///
///----------
/// FFI:
///----------
/// This API can be used in both trusted and untrusted partitions. See Freedom from Interference (FFI) concept for more details.
///
///------
///
///==================================================================		  			===================================================================================================
///Return value    								  									    Description
///==================================================================		  			===================================================================================================
///bds_outPwm_get_ts												                   The return structure containing;
///																							- Set current value in [mA]
///																							- Actual current measurement/current sensing of average of one PWM period in [mA]
///																							- Set value duty cycle in [permil]
///																							- Detailed diagnostic information OF the PWM output.
///																							- Function call status information (statusApi_e)
///
///==================================================================		   			===================================================================================================
///
///=======
///Code Example:
///=======
///============================================================================
///
/// PROGRAM appl_10ms_task
///
/// VAR
///
///     bds_outPwm_signal_e: bds_outPwm_signal_te; (* Declare the type for Pwm output signal*)
///
///     bds_outPwm_retGet_s: bds_outPwm_get_ts;    (* Declare the return structure of BDS-Function call*)
///
/// END_VAR
/// 
/// (* Initialize the signal value*)
///
/// bds_outPwm_signal_e := bds_outPwm_signal_te.bds_outPwm_K09_E;
/// 
/// (* Call BDS-Function to get the status of the output*)
///
/// bds_outPwm_retGet_s := bds_outPwm_get(bds_outPwm_signal_e);
/// 
/// (* Check return state of BDS-Function call*)
///
/// IF bds_outCmn_ok_E = bds_outPwm_retGet_s.statusApi_e THEN
///
///     (* Call successful, signal is valid*)
///
///     (* Status of output is updated successfully*)
///
/// ELSE
///
///     (* Handle error*)
///
/// END_IF;
///
/// END_PROGRAM
///
///============================================================================
{attribute 'external_name' := 'cmp_rts_bds_outPwm_get'}
FUNCTION bds_outPwm_get : bds_outPwm_get_ts
VAR_INPUT
	///The connector assigned signaVl name of the output.
	signal_e: USINT;
END_VAR

END_FUNCTION

// I/O API/OUT/API/bds_outPwm_cfgPeriod
///The BODAS API-function configures the period of a PWM high side or low side output in [us].
///
///=======
/// Remarks:
///=======
/// FOR the "low power low side outputs" the period range is FROM FROM 300us upto 31000us.

/// For the "high power high side outputs" the period range is from 1000us upto 100000us and for the "high power low side outputs" 4000us upto 100000us and only multiples of 1000us is configurable.

/// Default value of period is 10000us.
///
///----------
/// FFI:
///----------
/// This API can be used in trusted partitions. For untrusted partitions use bds_outPwm_cfgPeriod_ffi. See Freedom from Interference (FFI) concept for more details.
///
///------
///
///==================================================================		  			===================================================================================================
///Return value    								  									    Description
///==================================================================		  			===================================================================================================
///bds_outPwm_cfgPeriod_ts														            The return structure containing the state information (statusApi_e)
///
///==================================================================		   			===================================================================================================
///
///=======
///Code Example:
///=======
///============================================================================
///
/// PROGRAM appl_10ms_task
///
/// VAR
///
///     bds_outPwm_signal_e: bds_outPwm_signal_te; (* Define the structure of Pwm output signal*)
///
///     bds_outPwm_retCfgPeriod_s: bds_outPwm_cfgPeriod_ts; (* Declare return structure for the function call*)
///
///     tiPerd_us_u32: UDINT := 1000; (* Define the period in microseconds*)
///
/// END_VAR
/// 
/// (* Assign the Pwm signal type*)
///
/// bds_outPwm_signal_e := bds_outPwm_signal_te.bds_outPwm_K09_E;
/// 
/// (* Call function to configure the period of a Pwm output*)
///
/// bds_outPwm_retCfgPeriod_s := bds_outPwm_cfgPeriod(bds_outPwm_signal_e, tiPerd_us_u32);
/// 
/// (* Check return state of the BDS-Function call*)
///
/// IF bds_outCmn_ok_E = bds_outPwm_retCfgPeriod_s.statusApi_e THEN
///
///     (* If the call was successful and the signal is valid*)
///
///     (* The period of the Pwm output has been configured successfully*)
///
/// ELSE
///
///     (* Error handling*)
///
/// END_IF;
///
/// END_PROGRAM
///============================================================================
{attribute 'external_name' := 'cmp_rts_bds_outPwm_cfgPeriod'}
FUNCTION bds_outPwm_cfgPeriod : bds_outPwm_cfgPeriod_ts
VAR_INPUT
	///The connector assigned signal name of the output.
	signal_e: USINT;
	///The connector assigned signal name of the output.
	tiPerd_us_u32: UDINT;
END_VAR

END_FUNCTION

// I/O API/OUT/API/bds_outPwm_rstErr
/// The BODAS API-function reset the diagnostics error and unlocks the PWM high side or low side output.
///=======
/// Remarks:
///=======
/// +After a fault, the output is locked but the set point is still valid. With the reset OF the error the output is also unlocked.

/// +After a hot short circuit, the unlocking of the power output is only possible after a reactivation time of 2s.

/// +It is possible to poll the status of the fault. If the error has been healed, then the output can be reset.

/// +For over current fault: After reset, the output has to be switched on again using the API bds_outPwm_setDutyCycle or bds_outPwm_setCurrent.

/// +For more information see topic Proportional outputs.


///----------
/// FFI:
///----------
/// This API can be used in trusted partitions. For untrusted partitions use bds_outPwm_rstErr_ffi. See Freedom from Interference (FFI) concept for more details.
///
///
///==================================================================		  			===================================================================================================
///Return value    								  									    Description
///==================================================================		  			===================================================================================================
///bds_outPwm_rstErr_ts													                The return structure containing the state information (statusApi_e)
///
///==================================================================		   			===================================================================================================
///
///=======
///Code Example:
///=======
///============================================================================
/// PROGRAM appl_10ms_task
///
/// VAR
///
///     bds_outPwm_signal_e: bds_outPwm_signal_te; (* Define the structure of Pwm output signal*)
///
///     bds_outPwm_retRstErr_s: bds_outPwm_rstErr_ts; (* Declare return structure for the function call
///
/// END_VAR
/// 
/// (* Assign the Pwm signal type*)
///
/// bds_outPwm_signal_e := bds_outPwm_signal_te.bds_outPwm_K09_E;
/// 
/// (* Call function to reset the Pwm output diagnostic error and unlock the Pwm output*)
///
/// bds_outPwm_retRstErr_s := bds_outPwm_rstErr(bds_outPwm_signal_e);
/// 
/// (* Check return state of the BDS-Function call*)
///
/// IF bds_outCmn_ok_E = bds_outPwm_retRstErr_s.statusApi_e THEN
///
///     (* If the call was successful and the signal is valid*)
///
///     (* The diagnostic error for the output has been reset and the output is unlocked*)
///
/// ELSE
///
///     (* Error handling*)
///
/// END_IF;
///
/// END_PROGRAM
///
///============================================================================
{attribute 'external_name' := 'cmp_rts_bds_outPwm_rstErr'}
FUNCTION bds_outPwm_rstErr : bds_outPwm_rstErr_ts
VAR_INPUT
	///The connector assigned signal name of the output.
	signal_e: USINT;
END_VAR

END_FUNCTION

// I/O API/OUT/API/bds_outPwm_setCurrent
///The BODAS API-function sets the current for the PWM high side or low side output which is configured as closed loop current control mode.
///
///Set current range is from 0mA upto 3000mA/4000mA Current control upper limit depends on the used output, refer to RC27-18/40 - Outputs
///
///=======
/// Remarks:
///=======
///  + After a fault the output is locked but the set point is still valid.
///
///  + For more information see topic Proportional outputs.

///
///
///----------
/// FFI:
///----------
///This API can be used in trusted partitions . For untrusted partitions use |bds_out_do_getCurrent_ffi|. See Freedom from Interference (FFI) concept for more details.
///
///---------
/// Info
///---------
/// It is mandatory that the proportional output is configured as proportional output with closed loop current control mode, refer to bds_outPwm_cfgMode.

///---------
/// Attention
/// ---------
/// It is possible to poll the status of the fault. If the error has been healed, then the output can be unlocked by calling THIS API-FUNCTION.
///
/// After a hot short circuit and over current the unlock of the high power output is only possible after a reactivation wait time of 2s, refer to bit in status bds_outCmn_statusDiag_tb.

///==================================================================		  			===================================================================================================
///Return value    								  									    Description
///==================================================================		  			===================================================================================================
/// bds_outPwm_setCurrent_ts															The return structure containing the state information (statusApi_e)
///
///==================================================================		   			===================================================================================================
///
///=======
///Code Example:
///=======
///============================================================================
///
/// PROGRAM appl_10ms_task
///
/// VAR
///
///  bds_outPwm_signal_e: bds_outPwm_signal_te; (* Structure of PWM output signal*)
///
///  bds_outPwm_cfgMode_e: bds_outPwm_cfgMode_te; (* Output mode structure*)
///
///  bds_outPwm_retSetCurrent_s: bds_outPwm_setCurrent_ts; (* Return structure for setting current*)
///
///  bds_outPwm_set_i_mA_u16: UINT := 500; (* Define the set-current in mA*)
///
/// END_VAR
///
////// bds_outPwm_signal_e := bds_outPwm_signal_te.bds_outPwm_K09_E;
/// 
/// (* Configure the output as closed loop control mode*)
///
/// bds_outPwm_cfgMode(bds_outPwm_signal_e, bds_outPwm_cfgMode_e);
/// 
/// (* Actuate the PWM output with set-current*)
///
/// bds_outPwm_retSetCurrent_s := bds_outPwm_setCurrent(bds_outPwm_signal_e, bds_outPwm_set_i_mA_u16);
/// 
/// (* Check the return state of the BDS-Function call*)
///
/// IF bds_outCmn_ok_E = bds_outPwm_retSetCurrent_s.statusApi_e THEN
///
///     (* If the call was successful and the signal is valid*)
///
///     (* The PWM output has been actuated to the requested set-current successfully*)
///
/// ELSE
///
///     (* Error handling*)
///
/// END_IF;
///
/// END_PROGRAM
///============================================================================
{attribute 'external_name' := 'cmp_rts_bds_outPwm_setCurrent'}
FUNCTION bds_outPwm_setCurrent : bds_outPwm_setCurrent_ts
VAR_INPUT
	///The connector assigned signal name of the output.
	signal_e: USINT;
	///Storage address of the value.
	///
	///   defining the set current value for a PWM output which is configured as closed loop control current with the resolution in [mA]
	i_mA_u16: UINT;
END_VAR

END_FUNCTION

// I/O API/OUT/API/bds_outPwm_cfgMode
///The BODAS API-function configures the PWM high side or low side output as closed loop current control mode.
///
///=======
/// Remarks:
///=======
///With the closed loop current control mode further configurations are possible:
///
/// Software dither, refer to bds_outPwm_cfgDither.
///
/// Allowed current deviation from the set point, refer to bds_outPwm_cfgDiagCurrentDe.
///
/// Gain PI-Controller values for regulation (Kp and Ki), refer to bds_outPwm_cfgClc.



///
///----------
/// FFI:
///----------
/// This API can be used in both trusted and untrusted partitions. See Freedom from Interference (FFI) concept for more details.
///
///------
/// Info
///------
/// Only the proportional outputs with "Current Measurement" can be configured as closed loop current control mode which means output can be actuated with set-current.
///
/// Default output is in Pwm mode which means output can only be actuated with duty-cycle

///
///==================================================================		  			===================================================================================================
///Return value    								  									    Description
///==================================================================		  			===================================================================================================
///bds_outPwm_cfgMode_ts													            The return structure containing the state information (statusApi_e)
///
///==================================================================		   			===================================================================================================
///
///=======
///Code Example:
///=======
///============================================================================
///
///PROGRAM appl_10ms_task
///
///
///VAR
///
///    bds_outPwm_signal_e: bds_outPwm_signal_te; (* Declare and define the structure of Pwm output signal*)
///
///    bds_outPwm_cfgMode_e: bds_outPwm_cfgMode_te; (* Declare and define the output mode structure*)
///
///    bds_outPwm_retCfgMode_s: bds_outPwm_cfgMode_ts; (* Declare the return structure of BDS-Function call*)
///
///END_VAR
///
///(* Assign the Pwm signal type*)
///
///bds_outPwm_signal_e := bds_outPwm_signal_te.bds_outPwm_K09_E;
///
///(* Set the output mode to closed loop current control*)
///
///bds_outPwm_cfgMode_e := bds_outMode_CLCC_E;
///
///(* Call function to configure the output as closed loop current control mode*)
///
///bds_outPwm_retCfgMode_s := bds_outPwm_cfgMode(bds_outPwm_signal_e, bds_outPwm_cfgMode_e);
///
///(* Check return state of the BDS-Function call*)
///
///IF bds_outCmn_ok_E = bds_outPwm_retCfgMode_s.statusApi_e THEN
///
///    (* If the call was successful and the signal is valid*)
///
///    (* Output has been configured as closed loop current control successfully*)
///ELSE
///
///    (* Error handling*)
///
///END_IF;
///
/// END_PROGRAM
///============================================================================
{attribute 'external_name' := 'cmp_rts_bds_outPwm_cfgMode'}
FUNCTION bds_outPwm_cfgMode : bds_outPwm_cfgMode_ts
VAR_INPUT
	///The connector assigned signal name of the output.
	signal_e: USINT;
	///The connector assigned signal name of the output.
	mode_e: bds_outPwm_cfgMode_te;
END_VAR

END_FUNCTION

// I/O API/OUT/API/bds_outPwm_cfgDither
///The BODAS API-function configure the dither frequency and amplitude for the PWM high side or low side output which is configured as closed loop current control mode.
///
///=======
/// Remarks:
///=======
///   + The dither frequencies are predefined (see bds_outPwm_cfgDither_te) and its amplitude range is from 0 to 500mA.
///
///   + Default value for dither frequency is 0 [Hz] and amplitude is 0 [mA] (means dither configuration is disabled).
/// 
///----------
/// FFI:
///----------
///This API can be used in trusted partitions. For untrusted partitions use bds_outPwm_cfgDither_ffi. See Freedom from Interference (FFI) concept for more details.
///  
///------
/// Info:
///------
///
///The function is only possible for proportional outputs which has been configured as closed loop current control mode and a period of 1ms (f = 1000 Hz), refer to Outputs PWM  RC27-18/40 - Outputs
///
///==================================================================		  			===================================================================================================
///Return value    								  										 Description
///==================================================================		  			===================================================================================================
///bds_outPwm_cfgDither_ts																bds_outPwm_cfgDither_ts															
///
///==================================================================		   			===================================================================================================
///
///=======
///Code Example:
///=======
///============================================================================
///
/// PROGRAM appl_10ms_task 
///
/// VAR
///
///     bds_outPwm_signal_e: bds_outPwm_signal_te; (* Structure of PWM output signal*)
///
///     bds_outPwm_cfgMode_e: bds_outPwm_cfgMode_te; (* Output mode structure*)
///
///     bds_outPwm_cfg_ditherParams_s: bds_outPwm_ditherParams_ts; (* Structure for dither parameters.*)
///
///     bds_outPwm_retCfgDither_s: bds_outPwm_cfgDither_ts; (* Return structure for the dither configuration function*)
///
///     tiPerd_us_u32: UDINT := 1000; (* Define the period in microseconds
///
/// END_VAR
/// 
/// (* Set the PWM signal type*)
///
/// bds_outPwm_signal_e := bds_outPwm_signal_te.bds_outPwm_K09_E;
/// 
/// (* Configure the output as closed loop control mode*)
///
/// bds_outPwm_cfgMode(bds_outPwm_signal_e, bds_outPwm_cfgMode_e);
/// 
/// (* Set dither frequency and amplitude*)
///
/// bds_outPwm_cfg_ditherParams_s.ditherFrq_Hz_e := bds_outPwm_dither_90_Hz_E;
///
/// bds_outPwm_cfg_ditherParams_s.ditherAmp_mA_u16 := 400;
/// 
/// (* Configure the period for PWM output*)
///
/// bds_outPwm_cfgPeriod(bds_outPwm_signal_e, tiPerd_us_u32);
/// 
/// (* Configure the dither frequency and amplitude*)
///
/// bds_outPwm_retCfgDither_s := bds_outPwm_cfgDither(bds_outPwm_signal_e, bds_outPwm_cfg_ditherParams_s);
/// 
/// (* Check return state of the BDS-Function call*)
///
/// IF bds_outCmn_ok_E = bds_outPwm_retCfgDither_s.statusApi_e THEN
///
///     (* If the call was successful and the signal is valid,*)
///
///     (* The dither frequency and amplitude for the PWM output have been configured successfully*)
///
/// ELSE
///
///     (* Error handling*)
///
/// END_IF;
///
/// END_PROGRAM
///
///============================================================================
{attribute 'external_name' := 'cmp_rts_bds_outPwm_cfgDither'}
FUNCTION bds_outPwm_cfgDither : bds_outPwm_cfgDither_ts
VAR_INPUT
	///defining the output signal for the PWM output
	signal_e: USINT;
	///Frequency [Hz]
	///
	///   + defining the control structure values for the dither frequency and amplitude values of the selected PWM output which is configured as Closed Loop Control Current
	ditherParams_s: bds_outPwm_ditherParams_ts;
END_VAR

END_FUNCTION

// I/O API/OUT/API/bds_outPwm_cfgDiagCurrentDe
/// The BODAS API-function sets the current deviation for the PWM high side or low side output which is configured as closed loop current control mode.
/// 
///
///=======
/// Remarks:
///=======
///
/// Maximal allowed deviation between the set point AND the actual current is 500mA.
///
/// Value of 0mA deviation means the current deviation monitoring is disabled.
///
///If the value exceeds, the fault OR (out of range) is set after the debounce time elapses, but the output is not switched OFF.
///
/// If the deviation falls below the set deviation value, the fault OR is cleared after the debounce time elapses. 
///
/// For more information see bds_outPwm_get.


 
///----------
/// FFI:
///----------
///This API can be used in trusted partitions. For untrusted partitions use bds_outPwm_cfgDiagCurrentDe_ffi. See Freedom from Interference (FFI) concept for more details.
///
///
///==================================================================		  			===================================================================================================
///Return value    								  									    Description
///==================================================================		  			===================================================================================================
///bds_outPwm_cfgDiagCurrentDe_ts														The return structure containing the state information (statusApi_e)
///
///==================================================================		   			===================================================================================================
///
///=======
///Code Example:
///=======
///============================================================================
///
///PROGRAM appl_10ms_task
///
///VAR
///
///    bds_outPwm_signal_e: bds_outPwm_signal_te; (* Structure of PWM output signal*)
///
///    bds_outPwm_cfgMode_e: bds_outPwm_cfgMode_te; (* Output mode structure*)
///
///    bds_outPwm_retCfgDiagCurrentDe_s: bds_outPwm_cfgDiagCurrentDe_ts; (* Return structure for configuring current deviation*)
///
///    bds_outPwm_cfg_iDe_mA_u16: UINT := 300; (* Define the set-deviation in mA*)
///
/// END_VAR
///
/// bds_outPwm_signal_e := bds_outPwm_signal_te.bds_outPwm_K09_E;
///
///(* Configure the output as closed loop control mode*)
///
///bds_outPwm_cfgMode(bds_outPwm_signal_e, bds_outPwm_cfgMode_e);
///
///(* Call function to configure the current deviation*)
///
///bds_outPwm_retCfgDiagCurrentDe_s := bds_outPwm_cfgDiagCurrentDe(bds_outPwm_signal_e, bds_outPwm_cfg_iDe_mA_u16);
///
///(* Check the return state of the BDS-Function call*)
///
///IF bds_outCmn_ok_E = bds_outPwm_retCfgDiagCurrentDe_s.statusApi_e THEN
///
///    (* If the call was successful and the signal is valid*)
///
///    (* The current deviation for the PWM output has been configured successfully*)
///
///ELSE
///
///    (* Error handling*)
//
///END_IF;
///
/// END_PROGRAM
///============================================================================
{attribute 'external_name' := 'cmp_rts_bds_outPwm_cfgDiagCurrentDe'}
FUNCTION bds_outPwm_cfgDiagCurrentDe : bds_outPwm_cfgDiagCurrentDe_ts
VAR_INPUT
	///The connector assigned signal name of the output.
	signal_e: USINT;
	/// defining the deviation current value for a PWM output which is configured as closed loop control current with the resolution in [mA]
	iDe_mA_u16: UINT;
END_VAR

END_FUNCTION

// I/O API/OUT/API/bds_outPwm_cfgClc
///The BODAS API-function configure closed loop control gain for the PWM high side or low side output which is configured as closed loop current control mode.
///
///=======
/// Remarks:
///=======
///   +Range Kp factor [0...2000] and set default value is 100.
///
///	  +Range Ki factor [0...500] and set default value is 25.
///
///----------
/// FFI:
///----------
/// This API can be used in trusted partitions. For untrusted partitions use bds_outPwm_cfgClc_ffi. See Freedom from Interference (FFI) concept for more details.
///   
///==================================================================		  			===================================================================================================
///Return value    								  									     Description
///==================================================================		  			===================================================================================================
///bds_outPwm_cfgClc_ts																	The return structure containing the state information (statusApi_e)																		
///
///==================================================================		   			===================================================================================================
///
///=======
///Code Example:
///=======
///============================================================================
///
/// PROGRAM appl_10ms_task
///
/// VAR
///
///     bds_outClcC_signal_e: bds_outPwm_signal_te; (* Structure of PWM output signal*)
///
///     bds_outPwm_cfgMode_e: bds_outPwm_cfgMode_te; (* Output mode structure*)
///
///     bds_outPwm_cfg_clcParams_s: bds_outPwm_clcParams_ts; (* Structure for closed loop control gain*)
///
///     bds_outPwm_retCfgClc_s: bds_outPwm_cfgClc_ts; (* Return structure of BDS-Function call*)
///
/// END_VAR
/// 
/// (* Set the PWM signal type*)
///
/// bds_outClcC_signal_e := bds_outPwm_signal_te.bds_outPwm_K09_E;
/// 
/// (* Configure the output as closed loop control mode*)
///
/// bds_outPwm_cfgMode(bds_outClcC_signal_e, bds_outPwm_cfgMode_e);
/// 
/// (* Define the closed loop control gains*)
///
/// bds_outPwm_cfg_clcParams_s.Kp_u16 := 500; (* Proportional gain*)
///
/// bds_outPwm_cfg_clcParams_s.Ki_u16 := 300; (* Integral gain*)
/// 
/// (* Call function to configure closed loop control gain*)
///
/// bds_outPwm_retCfgClc_s := bds_outPwm_cfgClc(bds_outClcC_signal_e, bds_outPwm_cfg_clcParams_s);
/// 
/// (* Check the return state of the BDS-Function call*)
///
/// IF bds_outCmn_ok_E = bds_outPwm_retCfgClc_s.statusApi_e THEN
///
///     (* If the call was successful and the signal is valid*)
///
///     (* Closed loop control gain for the PWM output has been configured successfully*)
///
/// ELSE
///
///     (* Error handling*)
///
/// END_IF;
///
/// END_PROGRAM
///
///============================================================================
{attribute 'external_name' := 'cmp_rts_bds_outPwm_cfgClc'}
FUNCTION bds_outPwm_cfgClc : bds_outPwm_cfgClc_ts
VAR_INPUT
	///defining the output signal for the PWM output
	signal_e: USINT;
	///defining the control structure values for the gain proportional and integral values of the selected PWM output which is configured as Closed Loop Control Current
	///   + 0 to 500
	clcParams_s: bds_outPwm_clcParams_ts;
END_VAR

END_FUNCTION

// I/O API/OUT/API/bds_outPwm_cfgDiag
///The BODAS API-FUNCTION configures the diagnostic features FOR the PWM high side OR low side output.
///
/// Control the testpulses of PWM high power high side or low side output.
///
/// Control the PWM high side or low side output and also disabled its all diagnosis.
///
/// Control the non-hoterror short circuit detection of high side and low side PWM output.
///
/// Control the open load detection of PWM high side or low side output.
///
///=======
/// Remarks:
///=======
///
/// Control the testpulse OF PWM output:
///
/// Testpulses are enabled by default. Hence it can be disabled and enabled for the PWM high power high side or low side output.
///
///For example in some application the test pulses may disturb the required functionality of an output. For example if the high side PWM output is used as power supply for low power low side output.
///
///The testpulses can be enabled and disabled for High Power Outputs only.

///Attention 
///
///If testpulses are disabled for an output, fault detection and healing is limited. Please refer to topic Proportional outputs.

/// Control the PWM high side OR low side output AND disable its diagnosis:
///
/// Disable an unsed output and its diagnosis.
///
///The output should be disabled during start up of the application.

/// Attention
///
/// + Control the open load detection of high side and low side PWM output:
///  
/// + Open load detection is enabled by default. Hence it can be disabled and enabled for the PWM high side or low side output.
///  
/// + If open load detection is disabled, Open load will not be detected and healed.
///  
/// + For example in some application the open load detection may disturb the required functionality of an output. For example if the high power high side PWM output is used as power supply for the low side PWM output.
///  
/// + Please refer topic Proportional outputs for open load detection of PWM high side and low side output. 
///  
/// + Control the non-hot short circuit detection of high side and low side PWM output:
///  
/// + Non hot short circuit detection is enabled by default. Hence it can be disabled and enabled for the PWM high side or low side output.
///  
/// + If non hot short circuit detection is disabled, Non hot short circuit will not be detected and healed.
///  
/// + For high side PWM output short circuit to battery is non hot error and for low side PWM output short circuit to ground is non hot error.
///  
/// + Please refer topic Proportional outputs for non-hot short circuit detection of PWM high side and low side output. 


///----------
/// FFI:
///----------
/// This API can be used in trusted partitions. FOR untrusted partitions use bds_outPwm_cfgDiag_ffi. See Freedom FROM Interference (FFI) concept FOR more details.
///
///------
/// Info:
///------
/// Diagnostic configurations shall be disabled during start up of the application, otherwise faults may be detected on the time of diagnostic configuration. The previously detected faults can be reset with bds_outPwm_rstErr.

///==================================================================		  			===================================================================================================
///Return value    								  									    Description
///==================================================================		  			===================================================================================================
///bds_outPwm_cfgDiag_ts													             The return structure containing the state information (statusApi_e)
///
///==================================================================		   			===================================================================================================
///
///=======
///Code Example:
///=======
///============================================================================
///
/// PROGRAM OsIniProc
///
/// VAR
///
/// bds_outPwm_signal_e: bds_outPwm_signal_te;
///
/// bds_outPwm_retCfgDiag_s: bds_outPwm_cfgDiag_ts;
///
/// bds_outPwm_diagParam_s: bds_outCmn_diagParam_ts;

///END_VAR

///bds_outPwm_signal_e := bds_outPwm_signal_te.bds_outPwm_K09_E;

///bds_outPwm_diagParam_s.diFullDiag_l := FALSE;
///
///bds_outPwm_diagParam_s.diCntlAndDiag_l := TRUE;
///
///bds_outPwm_diagParam_s.diOpenLoadDetn_l := FALSE;
///
///bds_outPwm_diagParam_s.diNonHotSCDetn_l := FALSE;
///
///bds_outPwm_retCfgDiag_s := bds_outPwm_cfgDiag(bds_outPwm_signal_e, bds_outPwm_diagParam_s);
///
///IF bds_outCmn_ok_E = bds_outPwm_retCfgDiag_s.statusApi_e THEN
///
///    (* Call successful, signal is valid *)
///
///    (* Configured the diagnostic features for Pwm output successfully *)
///
///ELSE
///
/// (* error handling *)
///
/// END_IF;
///
/// END_PROGRAM
///============================================================================
{attribute 'external_name' := 'cmp_rts_bds_outPwm_cfgDiag'}
FUNCTION bds_outPwm_cfgDiag : bds_outPwm_cfgDiag_ts
VAR_INPUT
	///The connector assigned signal name of the output.
	signal_e: USINT;
	/// defining the control structure values for the control of the selected PWM output
	diagParam_s: bds_outCmn_diagParam_ts;
END_VAR

END_FUNCTION

// I/O API/OUT/API/bds_outClcU_cfgClc
/// The BODAS API-Function resets an existing diagnostic fault error and reactivating of voltage outputs, which are switched off due to an error detection.
///
/// FFI:
///----------
/// This API can be used in trusted partitions. For untrusted partitions use bds_outClcU_rstErr_ffi. See Freedom from Interference (FFI) concept for more details.
///   
///==================================================================		  			===================================================================================================
///Return value    								  									     Description
///==================================================================		  			===================================================================================================
/// bds_outClcU_rstErr_ts																	The return structure containing the state information (statusApi_e)																		
///
///==================================================================		   			===================================================================================================
///
///=======
///Code Example:
///=======
///============================================================================
///
/// PROGRAM appl_10ms_task
///
///VAR
///
///    bds_outClcU_signal_e: bds_outClcU_signal_te;
///	
///    bds_outClcU_retCfgClc_s: bds_outClcU_cfgClc_ts;
///	
///    clcParams_s: bds_outClcU_clcParams_ts;
///	
///END_VAR
///
///bds_outClcU_signal_e := bds_outClcU_signal_te.bds_outClcU_K25_E;
///
///(* set closed loop controler parameter set values *)
///
///clcParams_s.Kp_u16 := 200;
///
///clcParams_s.Ki_u16 := 50;
///
///(* call BDS-Function *)
///
///bds_outClcU_retCfgClc_s := bds_outClcU_cfgClc(bds_outClcU_signal_e, clcParams_s);
///
///(* check return state of BDS-Function call *)
///
///IF bds_outCmn_ok_E = bds_outClcU_retCfgClc_s.statusApi_e THEN
///
///    (* Call successful, signal is valid *)
///	
///    (* closed loop controler values Kp and Ki set correct for requested voltage output *)
///	
///ELSE
///
///    (* error handling *)
///	
///END_IF
///
/// END_PROGRAM
///
///============================================================================
{attribute 'external_name' := 'cmp_rts_bds_outClcU_cfgClc'}
FUNCTION bds_outClcU_cfgClc : bds_outClcU_cfgClc_ts
VAR_INPUT
	///defining the output signal for the PWM output
	signal_e: USINT;
	///defining the control structure values for the gain proportional and integral values of the selected PWM output which is configured as Closed Loop Control Current
	///   + 0 to 500
	clcParams_s: bds_outClcU_clcParams_ts;
END_VAR

END_FUNCTION

// I/O API/OUT_LEGACY/bds_out_po_unlock
///Unlocks proportional output if there is no error anymore.
///
///=======
/// Remarks:
///=======
///   + After a fault the output is locked but the set point is still valid. 
///   + It is possible to poll the status of the fault. If the error has been healed, then the output can be unlocked.
///   + After a hot short circuit and over current the unlock of the power output is only possible after a reactivation time of 2s.
///   + For over current fault: after unlocking the output has to be switched on again by the api, see: |bds_out_pod|, |bds_out_po|.
///
///----------
/// FFI:
///----------
///This API can be used in trusted partitions only. See Freedom from Interference (FFI) concept for more details.
///
///==================================================================		  			===================================================================================================
///Return value    								  									Description
///==================================================================		  			===================================================================================================
///16#0000																				No error, unlocked successfully.
///16#0001																				Error output was locked by the MO Module.
///16#0002																				Error reactivation time not elapsed.
///16#0004																				Error DFC_SCB is set.
///16#0008																				Error DFC_SCG is set
///16#0010																				Error DFC_OL is set
///16#0020																				Error DFC_OT is set
///16#0040																				Error DFC_OR is set
///16#0080																				Error OC is reset, output is unlocked
///16#8000																				Error signal out of range
///
///==================================================================		   			===================================================================================================
///
///=======
///Code Example:
///=======
///============================================================================
///
///PROGRAM appl_10ms_task
///
///VAR
///
///	return_u16: UINT := 16#00;
///
///END_VAR
///
///
///(* reset error of output K73 *)
///
///return_u16 = bds_out_po_unlock(bds_out_po_signal_te.K73);
///
///
///============================================================================
{attribute 'external_name' := 'cmp_rts_bds_out_po_unlock'}
FUNCTION bds_out_po_unlock : UINT
VAR_INPUT
	///The connector assigned signal name of the output.
	signal_e: UINT;
END_VAR

END_FUNCTION

// I/O API/IN/API/bds_inPha_get
///The bds_inPha_get API function provides measurement data of the phase between two input signals with same frequency.
///
///The phase measurement could be used to read two interdependent frequency signals to get the phase information of the signals and is based on the frequency measurement and therefore the requirements from the frequency measurement are also valid for the phase measurement.
///
///=======
/// Remarks:
///=======
///    + The phase measurement channel has to be configured in easyConfig. The phase measurement will be automatically configured during start up of the ECU.
///    + Certain input signals are grouped into predefined input pairs for phase measurement.
///    + For more information about the signal acquisition see Frequency aquisition.
///    + The measured phase shift between the primary and secondary input signal is given in [dDeg] and the range is defined from 0[dDeg] to +1800[dDeg] and -1800[dDeg] to 0[dDeg], reference is the rising edge of the primary signal.
///    + The measured phase difference between the primary and secondary input signal is given in [ns], reference is the rising edge of the primary signal.
///    + The measured phase period time of the primary and secondary input signal is given in [ns], range is defined from 50.000ns to 1.000.000.000ns (1Hz to 20kHz).
///    + The measured number of pulses of primary and secondary input signal is given with a 24-Bit counter with overflow (decimal range from 0 to 16.777.215). Pulses are counted with rising edge detection.
///    + The measured status information of the primary and secondary input signal is given as a bit field. There are error bits for maximum period overflow for primary and secondary signal and frequency mismatch.
///    + The maximum time for the period overflow detection of the primary and secondary signal is configured in easyConfig. There is only one time parameter for both signals.
///    + A frequency mismatch between primary and secondary signal is detected, if the time deviation between primary and secondary signal period is greater then 2000ns.
///    + A call of a configuration function is not required.
///    + If function is called with an invalid channel the function call status returns an error and all other values are set to "0"

///=======
/// Info:
///=======
///If a frequency mismatch is detected a status bit is set and for further diagnostic the phase measurement data for primary and secondary is still available (phase information should be used with caution).

///=======
/// Attention:
///=======
///If no input signal is present for some time and a signal is applied to the input pin, the first Api call returns a signal error information (bds_inPha_statusDiag_tb) and valid signal information is returned from the second Api call onwards. We recommend calling the API cyclically!

///
///----------
/// FFI:
///----------
///This API can be used in both trusted and untrusted partitions. See Freedom from Interference (FFI) concept for more details.
///	
///==================================================================		  			===================================================================================================
///Return value    								  									Description
///==================================================================		  			===================================================================================================
///|bds_inPha_measmt_ts|															The return structure containing the phase measurement values and state information for one measured sample
///
///==================================================================		   			===================================================================================================
///
///=======
///Code Example:
///=======
///============================================================================
///
///PROGRAM appl_10ms_task
///VAR bds_inPha_getMeasmPha_s: bds_inPha_measmt_ts;
/// appl_phaShift_dDeg_s32: INT;
/// appl_tiPhaDif_ns_u32: UDINT;
/// appl_tiPerdPrimSig_ns_u32: UDINT;
/// appl_tiPerdSecSig_ns_u32: UDINT;
/// appl_cntPlsPrimSig_u32: UDINT;
/// appl_cntPlsSecSig_u32: UDINT;
///END_VAR

///bds_inPha_getMeasmPha_s := bds_inPha_get(bds_inPha_K54_K37_E);
///IF bds_inCmn_ok_E = bds_inPha_getMeasmPha_s.status_e THEN
/// IF (0 = bds_inPha_getMeasmPha_s.statusDiag_b.stErrPrimSigMaxPerdOvf_b1) AND (0 = bds_inPha_getMeasmPha_s.statusDiag_b.stErrSecSigMaxPerdOvf_b1) AND (0 = bds_inPha_getMeasmPha_s.statusDiag_b.stErrSigFrqMismatch_b1) THEN
/// appl_phaShift_dDeg_s32 := bds_inPha_getMeasmPha_s.phaShift_dDeg_s32;
/// appl_tiPhaDif_ns_u32 := bds_inPha_getMeasmPha_s.tiPhaDif_ns_u32;
/// appl_tiPerdPrimSig_ns_u32 := bds_inPha_getMeasmPha_s.tiPerdPrimSig_ns_u32;
/// appl_tiPerdSecSig_ns_u32 := bds_inPha_getMeasmPha_s.tiPerdSecSig_ns_u32;
/// appl_cntPlsPrimSig_u32 := bds_inPha_getMeasmPha_s.cntPlsPrimSig_u32;
/// appl_cntPlsSecSig_u32 := bds_inPha_getMeasmPha_s.cntPlsSecSig_u32;
/// ELSE (* Error handling *)
/// END_IFELSE (* Error handling *)
///END_IF
///
///============================================================================
///
{attribute 'external_name' := 'cmp_rts_bds_inPha_get'}
FUNCTION bds_inPha_get : bds_inPha_measmt_ts
VAR_INPUT
	///The signal name that is assigned to the respective pin configured as current input
	signal_e: USINT;
END_VAR

END_FUNCTION

// I/O API/IN/API/bds_inPha_getTiBufd
///The bds_inPha_getTiBufd API function provides the phase measurement data of the last 20 periods. These samples can be used to perform an application specific filtering of the phase measurement data.
///
///=======
/// Remarks:
///=======
///    +The phase measurement channel has to be configured in easyConfig. The phase measurement will be automatically configured during start up of the ECU.
///	   +Specific frequency input signals are grouped into predefined input pairs for phase measurement.
///    +For more information about the signal acquisition see Frequency aquisition.
///    +The measured phase difference samples between the primary and secondary input signal is given in [ns], reference is the rising edge of the primary signal.
///    +The measured phase period time samples of the primary and secondary input signal is given in [ns], range is defined from 50.000ns to 1.000.000.000ns (1Hz to 20kHz).
///    +The measured number of pulses of primary and secondary input signal is given with a 24-Bit counter with overflow (decimal range from 0 to 16.777.215). Pulses are counted with rising edge detection.
///    +The measured number of newly received samples in the buffer since the last call of this API function is given from 0 to 20 samples.
///    +The measured status information of the primary and secondary input signal is given as a bit field. There are error bits for maximum period overflow for primary and secondary signal and frequency mismatch.
///    +The maximum time for the period overflow detection of the primary and secondary signal is configured in easyConfig. There is only one time for both signals.
///    +A frequency mismatch between primary and secondary signal is detected, if the time deviation between primary and secondary signal period is greater then 2000ns.
///    +A call of a configuration function is not required.

///=======
/// Info:
///=======
///If a frequency mismatch is detected a status bit is set and for further diagnostic the phase measurement data for primary and secondary is still available (phase information should be used with caution).

///=======
/// Attention:
///=======
///If no input signal is present for some time and a signal is applied to the input pin, the first Api call returns a signal error information (bds_inPha_statusDiag_tb) and valid signal information is returned from the second Api call onwards. We recommend calling the API cyclically!

///
///----------
/// FFI:
///----------
///This API can be used in both trusted and untrusted partitions. See Freedom from Interference (FFI) concept for more details.
///	
///==================================================================		  			===================================================================================================
///Return value    								  									Description
///==================================================================		  			===================================================================================================
///|bds_inPha_tiBufd_ts|															The return structure containing the status of the function call
///
///==================================================================		   			===================================================================================================
///
///=======
///Code Example:
///=======
///============================================================================
///
///PROGRAM appl_10ms_task
///
///VAR
///    bds_inPha_getTiBufd_s : bds_inPha_tiBufdMeasmt_ts;
///    bds_inPha_getTiBufdRet_s : bds_inPha_tiBufd_ts;
///
///    appl_tiPhaDif_ns_au32 : ARRAY [0..19] OF UINT;
///    appl_tiPerdPrimSig_ns_au32 : ARRAY [0..19] OF UINT;
///    appl_tiPerdSecSig_ns_au32 : ARRAY [0..19] OF UINT;
///    appl_cntPlsPrimSig_u32 : UINT;
///    appl_cntPlsSecSig_u32 : UINT;
///    appl_cntNewSample_u32 : UINT;
///    idxPhaSig_u8 : BYTE;
///
///    statusDiag_b : BOOL;  // Add a boolean for error handling logic
///END_VAR
///
/// Get the buffered phase between signal on pin K54 and on pin K37
///bds_inPha_getTiBufdRet_s := bds_inPha_getTiBufd(bds_inPha_K54_K37_E, bds_inPha_getTiBufd_s);
///
/// Check the returned status of the function call
///IF bds_inCmn_ok_E = bds_inPha_getTiBufdRet_s.status_e THEN
///
///    // Check the status of the signals
///    IF (NOT bds_inPha_getTiBufd_s.statusDiag_b.stErrPrimSigMaxPerdOvf_b1) AND
///       (NOT bds_inPha_getTiBufd_s.statusDiag_b.stErrSecSigMaxPerdOvf_b1) AND
///       (NOT bds_inPha_getTiBufd_s.statusDiag_b.stErrSigFrqMismatch_b1) THEN
///
///        // Copy the actual phase measurement times and counter into local variable
///        FOR idxPhaSig_u8 := 0 TO 19 DO
///            appl_tiPhaDif_ns_au32[idxPhaSig_u8] := bds_inPha_getTiBufd_s.tiPhaDif_ns_au32[idxPhaSig_u8];
///            appl_tiPerdPrimSig_ns_au32[idxPhaSig_u8] := bds_inPha_getTiBufd_s.tiPerdPrimSig_ns_au32[idxPhaSig_u8];
///            appl_tiPerdSecSig_ns_au32[idxPhaSig_u8] := bds_inPha_getTiBufd_s.tiPerdSecSig_ns_au32[idxPhaSig_u8];
///        END_FOR
///
///        appl_cntPlsPrimSig_u32 := bds_inPha_getTiBufd_s.cntPlsPrimSig_u32;
///        appl_cntPlsSecSig_u32 := bds_inPha_getTiBufd_s.cntPlsSecSig_u32;
///        appl_cntNewSample_u32 := bds_inPha_getTiBufd_s.cntNewSample_u32;
///
///    ELSE
///        // Error handling for signal status issues
///        statusDiag_b := TRUE;
///    END_IF
///
///ELSE
///    // Error handling for function call failure
///    statusDiag_b := TRUE;
///END_IF
///
///
///============================================================================
///
{attribute 'external_name' := 'cmp_rts_bds_inPha_getTiBufd'}
FUNCTION bds_inPha_getTiBufd : bds_inPha_tiBufd_ts
VAR_INPUT
	///The signal name that is assigned to the respective pin configured as current input
	signal_e: USINT;
	//The signal name that is assigned to the respective pin configured as current input
	tiBuf_ps: POINTER TO bds_inPha_tiBufdMeasmt_ts;
END_VAR

END_FUNCTION

// System API/DSM/DSM Refactored( 3-byte DTC)/API/bds_dsmDTC_getDTCVal
(*This function returns the DTC value of a specified DFC ID
=======
 Remarks:
=======
    -

----------
 FFI:
----------
This API can be used only in trusted partitions.  See Freedom from Interference (FFI) concept for more details.

==================================================================		  			===================================================================================================
Return value    								  									Description
==================================================================		  			===================================================================================================
|bds_dsmDTC_getDTCVal_ts|																The return structure containing the DTC value and API return status.
==================================================================		   			===================================================================================================


==================================================================		  			===================================================================================================
Possible status_e values for this function   								  		Description
==================================================================		  			===================================================================================================
bds_dsmCmn_ok_E																	    Call successful
bds_dsmCmn_outOfRng_E																The ID value passed as input to this API function is out of DFC ID ranges.
																					This is possible when the input ID passed to the API is passed as a numerical value instead of <DFC_Name>.id
==================================================================		   			===================================================================================================

=======
Code Example:
=======
============================================================================

PROGRAM appl_10ms_task
VAR

	appl_dsmDTC_getDTCVal_s: bds_dsmDTC_getDTCVal_ts ;
	dtcTest_u32 : UDINT;
	dfcId_u16 : UINT;

END_VAR

// Get DTC value of a given DFC 

appl_dsmDTC_getDTCVal_s := bds_dsmDTC_getDTCVal(dfcId_u16);

============================================================================

*)

(*This POU  returns the DTC value of a specified DFC ID.*)
{attribute 'external_name' := 'cmp_rts_bds_dsmDTC_getDTCVal'}
FUNCTION bds_dsmDTC_getDTCVal : bds_dsmDTC_getDTCVal_ts
VAR_INPUT
	(*Identifier corresponding to the DFC*)
	dfcId_u16 : UINT;
END_VAR

END_FUNCTION

// System API/DSM/DSM Refactored( 3-byte DTC)/API/bds_dsmDTC_updateErr
(*This function updates the DFES entry and the status of DTC, for faults with and without debouncing. It will set/heal the error with the help of DTC as input.
=======
 Remarks:
=======
    + Refer Diagnostic Debounce and Report Check on further details on how error debouncing works in BODAS-BSW.

----------
 FFI:
----------
This API can be usedin trusted partitions only.  See Freedom from Interference (FFI) concept for more details.

==================================================================		  			===================================================================================================
Return value    								  									Description
==================================================================		  			===================================================================================================
|bds_dsmDTC_updateErr_ts|															The return structure containing the return status of the function.
==================================================================		   			===================================================================================================


==================================================================		  			===================================================================================================
Possible status_e values for this function   								  		Description
==================================================================		  			===================================================================================================
bds_dsmCmn_ok_E																	    Call successful and DTC is set/healed. 
bds_dsmCmn_outOfRng_E																+ The input DTC value is present in neither ASW Errors nor BSW Errors.
																					+ fltLvl_e input is passed with values other than the enum values as in bds_dsmCmn_fltLvl_te

==================================================================		   			===================================================================================================

=======
Code Example:
=======
============================================================================

PROGRAM appl_10ms_task
VAR

	appl_updateErr_s: bds_dsmDTC_updateErr_ts ;
	fltLvl_e: bds_dsmCmn_fltLvl_te := bds_dsmCmn_fltLvl_100_Perc_e;
	tdiff_us_u32 : UDINT := 10000;

END_VAR

// Update the Error with 100% debounce active to make it Active Error 

appl_updateErr_s := bds_dsmDTC_updateErr(appl_dsmDTC_getDTCVal_s.dtc_u32, fltLvl_e, tdiff_us_u32);

============================================================================

*)
(*This POU is used to set a DTC to active / deactive based on the inputs provided.It updates the DFES entry, with the help of a DTC.*)
{attribute 'external_name' := 'cmp_rts_bds_dsmDTC_updateErr'}
FUNCTION bds_dsmDTC_updateErr : bds_dsmDTC_updateErr_ts
VAR_INPUT
	(*DTC Value*)
	dtc_u32 : UDINT;
	(*Fault level as result of the check (fault %)*)
	fltLvl_e : bds_dsmCmn_fltLvl_te;
	(*Time difference since last call in microseconds.*)
	tdiff_us_u32 : UDINT;	
END_VAR

END_FUNCTION

// System API/DSM/DSM Refactored( 3-byte DTC)/API/bds_dsmDTC_deleteErr
(*This function resets the status of specific DFC as well as deletes the related DFES entry if it exists through DTC.
=======
 Remarks:
=======
    -


----------
 FFI:
----------
This API can be used in trusted partitions only.  See Freedom from Interference (FFI) concept for more details.

==================================================================		  			===================================================================================================
Return value    								  									Description
==================================================================		  			===================================================================================================
|bds_dsmDTC_deleteErr_ts|																The return structure containing the return status of the API.

==================================================================		   			===================================================================================================


==================================================================		  			===================================================================================================
Possible status_e values for this function   								  		Description
==================================================================		  			===================================================================================================
bds_dsmCmn_ok_E																	    Call successful DTC status is reset and removed from DFES entry
bds_dsmCmn_outOfRng_E																The input DTC value is present in neither ASW Errors nor BSW Errors.
bds_dsmCmn_notAvl_E																	DTC is already cleared from DFES entry and status.
bds_dsmCmn_errInt_E																	Not available due to an internal error
==================================================================		   			===================================================================================================

=======
Code Example:
=======
============================================================================
PROGRAM appl_10ms_task
VAR
	appl_deleteErr_s: bds_dsmDTC_deleteErr_ts ;
	dtcTest_u32 : UDINT;

END_VAR

// Delete the error for the respective DTC value

appl_deleteErr_s := bds_dsmDTC_deleteErr(dtcTest_u32);

============================================================================

*)
(*This function resets the status of specific DFC as well as deletes the related DFES entry if it exists through DTC.*)
{attribute 'external_name' := 'cmp_rts_bds_dsmDTC_deleteErr'}
FUNCTION bds_dsmDTC_deleteErr : bds_dsmDTC_deleteErr_ts
VAR_INPUT
	(*The assigned DTC value.*)
	dtc_u32: UDINT;
END_VAR

END_FUNCTION

// System API/DSM/DSM Refactored( 3-byte DTC)/API/bds_dsmDTC_getErrList
(*This function provides the DTC list and total number of errors present in the DFES.
=======
 Remarks:
=======
    -
----------
 FFI:
----------
This API can be used only in trusted partitions.  See Freedom from Interference (FFI) concept for more details.

==================================================================		  			===================================================================================================
Return value    								  									Description
==================================================================		  			===================================================================================================
|bds_dsmDTC_getErrList_ts|															The return structure containing API status, DTC list and number of errors present in the list.
==================================================================		   			===================================================================================================


==================================================================		  			===================================================================================================
Possible status_e values for this function   								  		Description
==================================================================		  			===================================================================================================
bds_dsmCmn_ok_E																	    Call successful and DTC list along with number of DTCs is obtained.
bds_dsmCmn_invldPrm_E																Invalid mask_u16 value passed as input.
bds_dsmCmn_outOfRng_E																API is called when the query has already reached the maximum value of list of DFC status memory.
==================================================================		   			===================================================================================================

==================================================================		  			===================================================================================================
Possible mask_u16 values for this function   								  		Description
==================================================================		  			===================================================================================================
bds_dsmCmn_setActvErrMsk_DU16														Define for "DFC is active" mask as per status of DFC
bds_dsmCmn_tstdOnceMsk_DU16															DFC was tested at least once since start or reset as per DFC status.
bds_dsmCmn_setTstdOkMsk_DU16														DFC was at least once OK tested since start or reset according to status of DFC. 
bds_dsmCmn_setFailedClrMsk_DU16														Fault occured at least once since error was detected from memory, with respect to the status of DFC. 
==================================================================		   			===================================================================================================

==================================================================		  			===================================================================================================
Possible strtFromBgn_l values for this function   								  		Description
==================================================================		  			===================================================================================================
TRUE																					Query is started from the beginning of DTC status memory.
FALSE																					Query is continued with the next index where the last query was finished.
																						(This index is saved in BSW internally once in-depending on the parameter mask).
==================================================================		   			===================================================================================================
=======
Code Example:
=======
============================================================================

PROGRAM appl_10ms_task
VAR

	appl_errList_s: ARRAY[1..32] OF bds_dsmDTC_getErrList_ts; ;
	mask_u16 : UINT;
	strtFromBgn_l : TRUE;

END_VAR

   /// Query first 32 DTCs of Active Error Mask

  appl_errList_s[0] = bds_dsmDTC_getErrList(mask_u16, strtFromBgn_l);

 

  /// Query next 32 DTCs of Active Error Mask 

  appl_errList_s[1] = bds_dsmDTC_getErrList(mask_u16, FALSE);


============================================================================

*)(*This function is used to get all DTCs with the specified status.*)
{attribute 'external_name' := 'cmp_rts_bds_dsmDTC_getErrList'}
FUNCTION bds_dsmDTC_getErrList : bds_dsmDTC_getErrList_ts
VAR_INPUT
	(*The kind of error status can be specified in detail by means of this mask.*)
	mask_u16 : UINT;
	(*Query position start from beginning / end of previous query*)
	strtFromBgn_l : BOOL;
END_VAR

END_FUNCTION

// System API/DSM/DSM Refactored( 3-byte DTC)/API/bds_dsmDTC_getStatus
(*This function provides:

		1.Status of a DTC as in 16 bit status word of DFC.

		2.Tested State of a DTC (short status on whether the DTC is Active/Previously Active/Deactive).

=======
 Remarks:
=======
    -

----------
 FFI:
----------
This API can be usedin trusted partitions only.  See Freedom from Interference (FFI) concept for more details.

==================================================================		  			===================================================================================================
Return value    								  									Description
==================================================================		  			===================================================================================================
|bds_dsmDTC_getStatus_ts|															Return structure containing:
																						+ API status
																						+ Error Tested Status (Active/Previously Active/Deactive)
																						+ Descriptive status bitfield containing 16 bit status of DTC as in Diagnostic Fault Check.

==================================================================		   			===================================================================================================


==================================================================		  			===================================================================================================
Possible status_e values for this function   								  		Description
==================================================================		  			===================================================================================================
bds_dsmCmn_ok_E																	    Call successful.
bds_dsmCmn_outOfRng_E																The input DTC value is present in neither ASW Errors nor BSW Errors.
==================================================================		   			===================================================================================================

=======
Code Example:
=======
============================================================================

PROGRAM appl_10ms_task
VAR

	appl_dsmDTC_getStatus_s: bds_dsmDTC_getStatus_ts ;
	dtcTest_u32 : UDINT;

END_VAR

// Check status of DTC

appl_dsmDTC_getStatus_s := bds_dsmDTC_getStatus(dtcTest_u32);

============================================================================

*)
(*This POU is used to get the 16 bit status word of a DTC (which contains the detailed status of a DFC), and Error Status of corresponding DFC (Active / Previously Active / Deactive).*)
{attribute 'external_name' := 'cmp_rts_bds_dsmDTC_getStatus'}
FUNCTION bds_dsmDTC_getStatus : bds_dsmDTC_getStatus_ts
VAR_INPUT
	(*DTC value*)
	dtc_u32: UDINT;
END_VAR

END_FUNCTION

// System API/DSM/DSM Refactored( 3-byte DTC)/API/bds_dsmDTC_getDFES
(*This function is used to get DTC values and total number of errors present in DFES entry.
=======
 Remarks:
=======
    + On a maximum, 32 different DFES entries are possible. 
	+ Status Mask will take time (max. 10ms) to update in global mask so return status has to be monitored


----------
 FFI:
----------
This API can be used in trusted partitions only.  See Freedom from Interference (FFI) concept for more details.

==================================================================		  			===================================================================================================
Return value    								  									Description
==================================================================		  			===================================================================================================
|bds_dsmDTC_getDFES_ts|																Return structure of the API containing:

																							+ Status of API execution

																							+ List of DTC entries in DFES entry

																							+ Number of DTCs present in DFES entry

==================================================================		   			===================================================================================================


==================================================================		  			===================================================================================================
Possible status_e values for this function   								  		Description
==================================================================		  			===================================================================================================
bds_dsmCmn_ok_E																	    Call successful and DTC list along with number of DTCs is obtained.
bds_dsmCmn_outOfRng_E																API is called when the query has already reached the maximum value of DTC.
bds_dsmCmn_invldPrm_E																Invalid mask_u16 value passed as input.															
==================================================================		   			===================================================================================================
==================================================================		  			===================================================================================================
Possible mask_u16 values for this function   								  		Description
==================================================================		  			===================================================================================================
bds_dsmCmn_setActvErrMsk_DU16														Define for "DFC is active" mask as per status of DFC
bds_dsmCmn_tstdOnceMsk_DU16															DFC was tested at least once since start or reset as per DFC status.
bds_dsmCmn_setTstdOkMsk_DU16														DFC was at least once OK tested since start or reset according to status of DFC. 
bds_dsmCmn_setFailedClrMsk_DU16														Fault occured at least once since error was detected from memory, with respect to the status of DFC. 
==================================================================		   			===================================================================================================

=======
Code Example:
=======
============================================================================

PROGRAM appl_10ms_task
VAR

	appl_getDFES_s: bds_dsmDTC_deleteErr_ts ;
	mask_u16 : UINT;
	idx_u8 : USINT;
	dtcDFES_u32 :  ARRAY[1..32] OF UDINT;

END_VAR

// Store DFES entries 

appl_getDFES_s := bds_dsmDTC_getDFES(mask_u16);

FOR idx_u8 := 1 TO 32 BY 1  DO
	dtcDFES_u32[idx_u8] := appl_getDFES_s.dtcListDFES_au32[idx_u8];
END_FOR;

============================================================================

*)
(*This function is used to get DTC values and total number of errors present in DFES entry.*)
{attribute 'external_name' := 'cmp_rts_bds_dsmDTC_getDFES'}
FUNCTION bds_dsmDTC_getDFES : bds_dsmDTC_getDFES_ts
VAR_INPUT
	(*The kind of error status can be specified in detail by means of this mask.*)
	mask_u16 : UINT;
END_VAR

END_FUNCTION

// System API/DSM/DSM Refactored( 3-byte DTC)/API/bds_dsmJ1939_getJ1939DTC
(*This API function returns for a given DTC, the following J1939 related parameters:
	+ SPN
	+ FMI
	+ OC

and the following Lamp States:
	+ MIL
	+ RSL
	+ AWL
	+ PRL

=======
 Remarks:
=======
    -

----------
 FFI:
----------
This API can be usedin trusted partitions only.  See Freedom from Interference (FFI) concept for more details.

==================================================================		  			===================================================================================================
Return value    								  									Description
==================================================================		  			===================================================================================================
|bds_dsmDTC_getJ1939DTC_ts|															Return structure containing function return and
																					J1939 related parameters such as SPN, FMI, Lampstates (MIL, RSL, AWL, PRL) and Occurrence Counter.
==================================================================		   			===================================================================================================


==================================================================		  			===================================================================================================
Possible status_e values for this function   								  		Description
==================================================================		  			===================================================================================================
bds_dsmCmn_ok_E																	    Call successful.
bds_dsmCmn_outOfRng_E																The input DTC value is present in neither ASW Errors nor BSW Errors.
==================================================================		   			===================================================================================================

=======
Code Example:
=======
============================================================================

PROGRAM appl_10ms_task
VAR

	appl_dsmDTC_getJ1939DTC_s: bds_dsmDTC_getJ1939DTC_ts ;
	testDtc_u32 : UDINT;

END_VAR

// Get the J1939 parameters for the given J1939 DTC

appl_dsmDTC_getJ1939DTC_s := bds_dsmJ1939_getJ1939DTC(testDtc_u32);

============================================================================

*)
(*This function is used to read the J1939 specific DTC data (SPN, FMI, Lamp states and Occurrence Counter) for a given DTC.*)
{attribute 'external_name' := 'cmp_rts_bds_dsmJ1939_getJ1939DTC'}
FUNCTION bds_dsmJ1939_getJ1939DTC : bds_dsmJ1939_getJ1939DTC_ts
VAR_INPUT
	(*The assigned DTC value.*)
	dtc_u32 : UDINT;	
END_VAR

END_FUNCTION

// Diagnostics API/UDS/API/bds_uds_registerRoutineF001Callback
///This function will registers the callback for the routine control identifier F001.
///
///=======
/// Remarks:
///=======
///    + This is the mandatory API to be used for routine control identifier F001.
///	+ This is the common register API for routine control F000 for all sub functions like start(), stop(), getResults().
///    + The |GVL_uds| is given for usage of defines.
///
///----------
/// FFI:
///----------
///This API can be used in trusted partitions only. See Freedom from Interference (FFI) concept for more details.
///
///==================================================================		  			===================================================================================================
///Return value    								  									Description
///==================================================================		  			===================================================================================================
///0																					No error
///1																					Invalid pointer
///
///==================================================================		   			===================================================================================================
///
///=======
///Code Example:
///=======
///============================================================================
///
///FUNCTION POU_3 : BYTE
///VAR_INPUT
///
///    dataIn1 : BYTE;
///
///    status : BYTE;
///
///    dataOut1 : POINTER TO BYTE;
///
///    Error_Code : POINTER TO BYTE;
///
///    subservice_u8 : BYTE;
///END_VAR
///
///VAR
///    data_au8: ARRAY[0..7] OF BYTE :=[1,2,3,4,5,6,7,8];
///
///    i: BYTE;
///
///    RidValue_u16: UINT;
///
///    set: BYTE;
///END_VAR
///
///IF(subservice_u8=1)
///
///    THEN bds_uds_setCallbackStatus(0);
///
///END_IF
///
///IF(subservice_u8=2)
///
///    THEN bds_uds_setCallbackStatus(0);
///
///END_IF
///
///IF(subservice_u8=3)
///
///    THEN bds_uds_setCallbackStatus(1);
///
///END_IF
///
///(*Registering callback*)
///
///PROGRAM POU_10
///VAR
///   
///    flag_3 : BOOL := 1;    
///
///END_VAR
///
///
///IF ( flag_3)
///
///    THEN bds_uds_registerRoutineF001Callback (ADR(POU_3));
///
///    flag_3 := 0;(*To make api call once in application*)
///
///END_IF
///
///
///============================================================================
{attribute 'external_name' := 'cmp_rts_bds_uds_registerRoutineF001Callback'}
FUNCTION bds_uds_registerRoutineF001Callback : USINT
VAR_INPUT
	///Function pointer with argument of as mentioned above
	func_pf: POINTER TO BOOL;
END_VAR

END_FUNCTION

// Communication API/CAN/CAN-FD legacy/API/bds_can_fd_getData
///Get the oldest message (FIFO) from the CAN-FD receive buffer of the specified CAN channel.
///
///=======
/// Remarks:
///=======
/// + A CAN-FD receive buffer is not available until a buffer is registered. For registering a buffer please refer How to configure CAN FD related parameters and related pages.
/// + First check the return value before accessing the message.
/// + The header file bds_cmn_bsw.h is included for enabling usage of defines. 
/// + For receiving CAN 2.0 messages refer bds_can_getData.
///
///----------
/// FFI:
///----------
///This API can be used in trusted partitions.
///
///==================================================================		  			===================================================================================================
///Return value    								  										Description
///==================================================================		  			===================================================================================================
///0 : bds_can_fd_ok_E																	Function is called without errors. Message data returned in msg_s are valid.
///14 : bds_can_fd_invldChnl_E															Invalid CAN channel.
///30 : bds_can_fd_rxBufOvfl_E															Receive buffer overflow. At least one message is lost. Message data returned in msg_s are valid.
///31 : bds_can_fd_rxBufEmpty_E															Receive buffer is empty. Message data returned in msg_s are invalid.
///32 : bds_can_fd_rxBufLenZero_E														Receive buffer length is zero. Message data returned in msg_s are invalid.
///60 : bds_can_fd_invldAddr_E															Invalid address (parameter msg_s).
///100 : bds_can_fd_paramChnl3Err_E														CAN-FD not supported in CAN_3.
///
///==================================================================		   			===================================================================================================
///
///=======
///Code Example:
///=======
///============================================================================
///PROGRAM appl_Task_1
///  VAR
///     msg_s: bds_can_Message_ts;
///  END_VAR
///
///  IF (0 = bds_can_getData(BDS_CAN_1_D, ADR(msg_s))) THEN
///  
///    (* Message in structure msg_s is valid and can be evaluated. *)
///	
///  END_IF
///END
///============================================================================

{attribute 'external_name' := 'cmp_rts_bds_can_fd_getData'}
FUNCTION bds_can_fd_getData : bds_can_fd_St_te
VAR_INPUT
	//Indicates the CAN channel.
	//Possible values :
	//BDS_CAN_1_D(0)
	//BDS_CAN_2_D(1)
	//BDS_CAN_4_D(3)
	chnl_e:bds_can_Chnl_te;
	//Pointer to the message data of type bds_can_fd_Message_ts.
	msg_s: POINTER TO bds_can_fd_Message_ts;
END_VAR

END_FUNCTION

// Communication API/CAN/CAN-FD legacy/API/bds_can_fd_getRxBufStatus
///This function returns the status of the CAN-FD receive buffer.
///
///=======
/// Remarks:
///=======
///  + The header file bds_cmn_bsw.h is included for enabling usage of defines.
/// 
///----------
/// FFI:
///----------
///This API can be used in trusted partitions.
///
///==================================================================		  			===================================================================================================
///Return value    								  										Description
///==================================================================		  			===================================================================================================
/// > 0																					Number of CAN messages in Rx buffer of the specified CAN channel which have been received.
///  0																					Rx buffer is empty.
/// -1																					Invalid CAN channel / CAN-FD not supported in CAN_3.
/// 
///
///==================================================================		   			===================================================================================================
///
///=======
///Code Example:
///=======
///============================================================================
///PROGRAM appl_Task_1
///  VAR
///    numMsg_s32: DINT := 16#00;
///  END_VAR
/// 
///  numMsg_s32 := bds_can_fd_getRxBufStatus(BDS_CAN_1_D);
///
///  IF (numMsg_s32 > 0) THEN
///  
///    (* RX buffer contains messages which can be read with bds_can_getData() *)
///	
///  END_IF
///END
///============================================================================
{attribute 'external_name' := 'cmp_rts_bds_can_fd_getRxBufStatus'}
FUNCTION bds_can_fd_getRxBufStatus : DINT

VAR_INPUT
	//Indicates the CAN channel.
	//Possible values :
	// + BDS_CAN_1_D(0)
	// + BDS_CAN_2_D(1)
	// + BDS_CAN_4_D(3)
	chnl_e:bds_can_Chnl_te;
END_VAR

END_FUNCTION

// Communication API/CAN/CAN-FD legacy/API/bds_can_fd_getTxBufStatus
///This function returns the status of the CAN-FD transmit buffer of a CAN channel.
///=======
/// Remarks:
///=======
/// + Status = number of CAN-FD messages in CAN-FD transmit buffer which have to be sent.
/// + The header file bds_cmn_bsw.h is included for enabling usage of defines.
///
///----------
/// FFI:
///----------
///This API can be used in trusted partitions.
///
///==================================================================		  			===================================================================================================
///Return value    								  										Description
///==================================================================		  			===================================================================================================
/// > 0																					Number of CAN-FD messages in CAN-FD transmit buffer of the specified CAN channel which have to be sent.
///	  0																					Tx buffer is empty.
/// - 1																					Invalid CAN channel / CAN-FD not supported in CAN_3.
///
///==================================================================		   			===================================================================================================
///
///=======
///Code Example:
///=======
///============================================================================
///PROGRAM appl_Task_1
///  VAR
///  
///    numMsg_s32: DINT := 16#00;
///  END_VAR
/// 
///  numMsg_s32 := bds_can_fd_getTxBufStatus(BDS_CAN_1_D);
/// 
///  IF (numMsg_s32 > 0) THEN
///  
///    (* TX buffer contains still messages which could not be sent. If CAN channel
///       is in operational mode the messages will be sent as soon as possible. *)
///	   
///  END_IF
///END
///============================================================================

{attribute 'external_name' := 'cmp_rts_bds_can_fd_getTxBufStatus'}

FUNCTION bds_can_fd_getTxBufStatus : DINT
VAR_INPUT
	//Indicates the CAN channel.
	//Possible values :
	//BDS_CAN_1_D(0)
	//BDS_CAN_2_D(1)
	//BDS_CAN_4_D(3)
	chnl_e: bds_can_Chnl_te;
END_VAR

END_FUNCTION

// Communication API/CAN/CAN-FD legacy/API/bds_can_fd_isTxChannelFree
///This function checks whether a complete CAN transmit channel is empty.
///
///=======
/// Remarks:
///=======
/// + Empty means that there is no message to send in hardware CAN controller and CAN-FD transmit buffer (if registered) is empty.
/// + This function can be used in order to check if a previous CAN-FD message was sent completely on CAN bus.
/// + The header file bds_cmn_bsw.h is included for enabling usage of defines.
///----------
/// FFI:
///----------
///This API can be used in trusted partitions.
///
///==================================================================		  			===================================================================================================
///Return value    								  										Description
///==================================================================		  			===================================================================================================
/// 0																					No error. CAN transmit channel is empty. No CAN message has to be sent at the moment. 
/// 1																					No error. CAN transmit channel is not empty. Sending of a message is still in progress and/or CAN Tx messages are still buffered for sending. 
/// 2																					Unknown CAN channel / CAN-FD not supported in CAN_3.
///==================================================================		   			===================================================================================================
///
///=======
///Code Example:
///=======
///============================================================================
///PROGRAM appl_Task_1
///  VAR
///  
///  END_VAR
///
///  IF (BDS_CAN_FD_TX_CHANNEL_EMPTY_DU16 = bds_can_fd_isTxChannelFree(BDS_CAN_1_D)) THEN
///  
///    (* All TX databoxes and TX buffer on CAN channel 1 are empty. *)
///    (* ... *)
///	
///  END_IF
///END
{attribute 'external_name' := 'cmp_rts_bds_can_fd_isTxChannelFree'}

FUNCTION bds_can_fd_isTxChannelFree : UINT
VAR_INPUT
	//Indicates the CAN channel.
	//Possible values :
	//BDS_CAN_1_D(0)
	//BDS_CAN_2_D(1)
	//BDS_CAN_4_D(3)
	chnl_e: bds_can_Chnl_te;
END_VAR

END_FUNCTION

// Communication API/CAN/CAN-FD legacy/API/bds_can_fd_registerRxBuf
///This API registers a CAN-FD transmit buffer for receiving data on a node.
///
///=======
/// Remarks:
///=======
/// + The header file bds_cmn_bsw.h is included for enabling usage of defines.
/// + This function must be called only in ASW Initialization task if required. Alternatively we can configure CAN-FD transmit buffer in easyConfig till value of 50 for a given CAN channel.
/// + Refer chapter How to configure CAN FD related parameters on a detailed note on how to configure CAN-FD buffers.
///----------
/// FFI:
///----------
///This API can be used in trusted partitions.
///
///==================================================================		  			===================================================================================================
///Return value    								  										Description
///==================================================================		  			===================================================================================================
///0 : bds_can_fd_ok_E																	Function is called without errors. Callback function was initialized successfully.			
///55 : bds_can_fd_ovlpAddr_E															New buffer overlaps current buffer.
///60 : bds_can_fd_invldAddr_E															address passed in argument buf_pas is Invalid
///18 : bds_can_fd_numMsgZero_E															Number of messages to be registered is zero
///99 : bds_can_fd_cfgNotAllowed_E														Configuration not allowed apart from ASW initialization task.
///100 : bds_can_fd_paramChnl3Err_E														CAN-FD not supported in CAN_3
///
///==================================================================		   			===================================================================================================
///=======
///Code Example:
///=======
///============================================================================
///PROGRAM PLC_PRG
/// VAR
///
/// rbr_can1_fd_rx_buf_as: ARRAY[1..10] OF bds_can_fd_Message_ts;
///
/// BDS_CANFD_NUM_OF_MESSAGES:UINT:=10;
///
/// flag: BOOL;
/// END_VAR
///
///
/// IF flag=FALSE THEN
///	bds_can_fd_registerRxBuf(BDS_CAN_1_D, ADR(rbr_can1_fd_rx_buf_as), BDS_CANFD_NUM_OF_MESSAGES);
///	flag:=TRUE;
/// END_IF
///END 
///============================================================================
{attribute 'external_name' := 'cmp_rts_bds_can_fd_registerRxBuf'}

FUNCTION bds_can_fd_registerRxBuf : bds_can_fd_St_te
VAR_INPUT
	//Indicates the CAN channel.
	//Possible values :
	//BDS_CAN_1_D(0)
	//BDS_CAN_2_D(1)
	//BDS_CAN_4_D(3)
	chnl_e:bds_can_Chnl_te;
	//Start address of CAN-FD receive buffer
	buf_pas: POINTER TO bds_can_fd_Message_ts;
	//Number of messages
	numMsg_u16: UINT;
END_VAR

END_FUNCTION

// Communication API/CAN/CAN-FD legacy/API/bds_can_fd_registerTxBuf
///This API registers a CAN-FD transmit buffer for transmitting data on a node.
///
///=======
/// Remarks:
///=======
/// + The header file bds_cmn_bsw.h is included for enabling usage of defines.
/// + This function must be called only in ASW Initialization task if required. Alternatively we can configure CAN-FD receive buffer in easyConfig (upto 50 buffers) for a given CAN channel.
/// + Refer chapter How to configure CAN FD related parameters on a detailed note on how to configure CAN-FD buffers.
///----------
/// FFI:
///----------
///This API can be used in trusted partitions.
///
///==================================================================		  			===================================================================================================
///Return value    								  										Description
///==================================================================		  			===================================================================================================
///0 : bds_can_fd_ok_E																	Function is called without errors. Callback function was initialized successfully.
///55 : bds_can_fd_ovlpAddr_E															New buffer overlaps current buffer.
///60 : bds_can_fd_invldAddr_E															Invalid address
///18 : bds_can_fd_numMsgZero_E															Number of messages to be registered is zero
///99 : bds_can_fd_cfgNotAllowed_E														Configuration not allowed apart from ASW Initialization task.
///100 : bds_can_fd_paramChnl3Err_E														CAN-FD not supported in CAN_3
///==================================================================		   			===================================================================================================
///
///=======
///Code Example:
///=======
///============================================================================
///PROGRAM PLC_PRG
/// VAR
///
/// rbr_can1_fd_tx_buf_as: ARRAY[1..10] OF bds_can_fd_Message_ts;
///
/// BDS_CANFD_NUM_OF_MESSAGES:UINT:=10;
///
/// flag: BOOL;
/// END_VAR
///
///
/// IF flag=FALSE THEN
///	bds_can_fd_registerTxBuf(BDS_CAN_1_D, ADR(rbr_can1_fd_tx_buf_as), BDS_CANFD_NUM_OF_MESSAGES);
///	flag:=TRUE;
/// END_IF
///END
///============================================================================
{attribute 'external_name' := 'cmp_rts_bds_can_fd_registerTxBuf'}

FUNCTION bds_can_fd_registerTxBuf : bds_can_fd_St_te
VAR_INPUT
	//Indicates the CAN channel.
	//Possible values :
	// + BDS_CAN_1_D(0)
	// + BDS_CAN_2_D(1)
	// + BDS_CAN_4_D(3)
	chnl_e:bds_can_Chnl_te;
	//Start address of CAN-FD transmit buffe 
	buf_pas: POINTER TO bds_can_fd_Message_ts;
	//Number of messages
	numMsg_u16: UINT;
END_VAR

END_FUNCTION

// Communication API/CAN/CAN-FD legacy/API/bds_can_fd_resetTxBuf
///This function resets the specified CAN-FD transmit buffer for a specified CAN channel.
///
///=======
/// Remarks:
///=======
/// + The header file bds_cmn_bsw.h is included for enabling usage of defines.
///
///----------
/// FFI:
///----------
///This API can be used in trusted partitions.
///
///
///==================================================================		  			===================================================================================================
///Return value    								  										Description
///==================================================================		  			===================================================================================================
/// 0																					Function is called without errors. CAN-FD Transmit buffer is reset.																	
/// 1																					Invalid buffer type. 
/// 3																					Unknown CAN channel.
/// 100																				    CAN-FD not supported in CAN_3.																			
///==================================================================		   			===================================================================================================
///
///=======
///Code Example:
///=======
///============================================================================
///
///PROGRAM appl_Task_1
///  VAR
///  
///  END_VAR
///
///  (* Tx buffer and all Tx data boxes of CAN channel 1 will be reset *)
///  
///  bds_can_fd_resetTxBuf(BDS_CAN_1_D, BDS_CAN_BUFTYPE_BUF_DU8 OR BDS_CAN_BUFTYPE_DATABOXES_DU8);
///
///  (* ... *)
///END
///
///============================================================================
{attribute 'external_name' := 'cmp_rts_bds_can_fd_resetTxBuf'}
FUNCTION bds_can_fd_resetTxBuf : UINT
VAR_INPUT
	//Indicates the CAN channel.
	//Possible values :
	// + BDS_CAN_1_D(0)
	// + BDS_CAN_2_D(1)
	// + BDS_CAN_4_D(3)
	chnl_e:bds_can_Chnl_te;
	//Indicates the buffer type:
	//Value 0 - No reset
	//Value 1 - BDS_CAN_BUFTYPE_BUF_DU8 - Reset CAN-FD Transmit Buffer
	bufType_u8: USINT;
END_VAR

END_FUNCTION

// Communication API/CAN/CAN-FD legacy/API/bds_can_fd_sendData
///Sends a CAN-FD message via the specified CAN channel.
///
///=======
/// Remarks:
///=======
/// + The CAN channel is not buffered until a buffer is registered. For registering a buffer please refer How to configure CAN FD related parameters and related pages.
/// + CAN-FD messages sent with this function is supported with BRS enabled only.
/// + If a CAN-FD transmit buffer is registered then messages are saved in buffer and will be sent in a background process as fast as possible. The buffer principle is first in first out (FIFO)..
/// + The header file bds_cmn_bsw.h is included for enabling usage of defines.
/// + For sending CAN 2.0 messages refer bds_can_sendData.
///----------
/// FFI:
///----------
///This API can be used in trusted partitions.
///
///==================================================================		  			===================================================================================================
///Return value    								  										Description
///==================================================================		  			===================================================================================================
///0 : bds_can_fd_ok_E																	Function is called without errors. CAN message will be sent.
///14 : bds_can_fd_invldChnl_E															Unknown CAN channel. 																				
///15 : bds_can_fd_invldId_E															Invalid CAN identifier.
///16 : bds_can_fd_invldFormat_E														Invalid message format.	
///17 : bds_can_fd_invldNumBytes_E														Invalid number of data bytes.
///20 : bds_can_fd_txBufOvfl_E															CAN message could not be sent, because of send buffer is full. *1)
///60 : bds_can_fd_invldAddr_E															Invalid address (parameter data_pau8).
///100 - bds_can_fd_paramChnl3Err_E														CAN-FD not supported in CAN_3.
///
///=======
///Code Example:
///=======
///============================================================================
///
///PROGRAM PLC_PRG
///  VAR
///  
///  END_VAR
///
///  (* remark: a CAN TX buffer must be configured in easyConfig *)
///
///  (* re-initialize can channel 1 with 250KBaud. Call the bds_can_init API once *)
///  
///  bds_can_init(BDS_CAN_1_D, BDS_BAUD_250K_DU32);
///
///  (* ... *)
///  
///END
///
///PROGRAM appl_Task_1
///  VAR
///    data_au8: ARRAY[0..63] OF USINT;
///  END_VAR
///
///  data_au8[0] := 5;
///  data_au8[1] := 7;
///
///  IF (0 = bds_can_fd_sendData(BDS_CAN_1_D, 16#123456, BDS_CAN_EXD_DU8, 2, ADR(data_au8))) THEN
///  
///    (* ok, message is buffered and will be sent as fast as possible. *)
///	
///  END_IF
///END
///============================================================================										
{attribute 'external_name' := 'cmp_rts_bds_can_fd_sendData'}

FUNCTION bds_can_fd_sendData : bds_can_fd_St_te
VAR_INPUT
	//Indicates the CAN channel.
	//Possible values :
	// + BDS_CAN_1_D(0)
	// + BDS_CAN_2_D(1)
	// + BDS_CAN_4_D(3)
	chnl_e: bds_can_Chnl_te; 
    //Identifier of CAN-FD message.
	//Value range:
	//0x000 .. 0x7FF (11-bit standard format .. 0x1FFFFFFF (29-BIT extented format
	id_u32: UDINT;
	//Indicates the format of the CAN-FD message.
	//Value range:
	//BDS_CAN_STD_DU8  (11-bit standard format)
	//BDS_CAN_EXD_DU8  (29-bit extented format)
 	format_u8 : USINT;
	//Number of bytes to be sent.
	//
	//Value range: 1 .. 64
	numBytes_u8: USINT;
	//Pointer to array of data bytes. The number of bytes is contained in parameter numBytes_u8.
	//A NULL pointer is allowed if number of data bytes (parameter numBytes_u8) is zero. 
	data_pau8: POINTER TO USINT;
END_VAR

END_FUNCTION

